SUBAPPLICATION Uebung_094b3c_AX (* Wie Uebung_094b3_AX, aber K=2 aktiviert zwei Optionsgruppen NACHEINANDER statt nur einer: OptionalGroup_001a wird vom DEMUX aktiviert und reicht die Aktivierung ueber ihren Plug PLUG1 an OptionalGroup_001b weiter - der DEMUX bekommt seine Bestaetigung erst, wenn BEIDE Gruppen initialisiert sind. *)
  (* Standard: 61499-2; Description: Copyright (c) 2026 Meisterschulen am Ostbahnhof This program and the accompanying materials are made available under the terms of the Eclipse Public License 2.0 which is available at https://www.eclipse.org/legal/epl-2.0/ SPDX-License-Identifier: EPL-2.0 *)
  (* Version 1.0, 2026-10-13, Franz Höpfinger, Meisterschulen am Ostbahnhof, Daisy-Chain-Variante von Uebung_094b3_AX: OptionalGroup_001 durch OptionalGroup_001a (mit zusaetzlichem Plug PLUG1) ersetzt und mit einer neuen OptionalGroup_001b dahinter verkettet - zeigt, wie man ueber die Plug/Socket-Kette mehrere Gruppen sequenziell (nacheinander, nicht gleichzeitig) hochfahren kann, ohne das Busy-Gating des DEMUX zu verletzen. *)
  PACKAGE Uebungen;
  IMPORT Uebungen::const::UT::DefaultPool::InputNumber_I1;
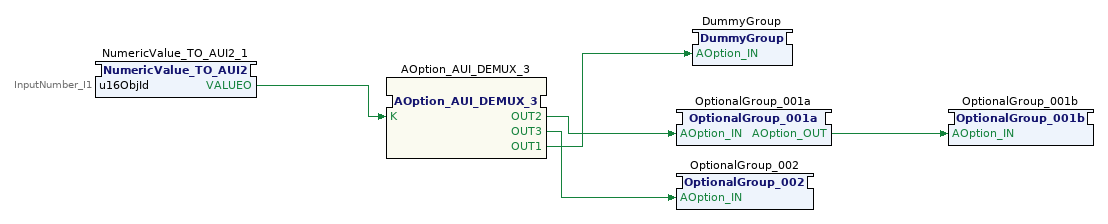
  FBS
    AOption_AUI_DEMUX_3 : Option::selection::AOption_AUI_DEMUX_3;
  END_FBS
  SUBAPPS
    NumericValue_TO_AUI2_1 : MyLib::sys::NumericValue_TO_AUI2(u16ObjId := InputNumber_I1);
    OptionalGroup_001a : MyLib_AX_Option::sys::OptionalGroup_001a;
    OptionalGroup_002 : MyLib_AX_Option::sys::OptionalGroup_002;
    DummyGroup : MyLib_AX_Option::sys::DummyGroup;
    OptionalGroup_001b : MyLib_AX_Option::sys::OptionalGroup_001b;
  END_SUBAPPS
  ADAPTER_CONNECTIONS
    NumericValue_TO_AUI2_1.VALUEO TO AOption_AUI_DEMUX_3.K;
    AOption_AUI_DEMUX_3.OUT2 TO OptionalGroup_001a.AOption_IN;
    AOption_AUI_DEMUX_3.OUT3 TO OptionalGroup_002.AOption_IN;
    AOption_AUI_DEMUX_3.OUT1 TO DummyGroup.AOption_IN;
    OptionalGroup_001a.AOption_OUT TO OptionalGroup_001b.AOption_IN;
  END_CONNECTIONS
END_SUBAPPLICATION
